(* IEC 61131-3 sources: SRCI_CLIENT_PLC/RobotLibrary/Library/Structures/AxesGroup/State/SyncState, 4 files *)

(* ---- AxesGroupStateSyncState.st ---- *)
{attribute 'pack_mode' := '1'}
// -------------------------------------------------------------------------
//  SRCI Robot Library
// -------------------------------------------------------------------------
//
//  Object:      AxesGroupStateSyncState
//  Author:      Thorsten Brach
//  Date:        2024-06-01
//
//  Description:
//
//
//  Copyright:
//    (C) 2024 Thorsten Brach. All rights reserved
//             Licensed under the MIT License.
//
//  Disclaimer:
//    This project is provided without any guarantee and can be used for
//    private and commercial purposes. Any use is at the user’s
//    own risk and responsibility.
//
// -------------------------------------------------------------------------
TYPE AxesGroupStateSyncState :
STRUCT
  /// Bit 00: Tool
  Tool             : BOOL;
  /// Bit 01: Frame
  Frame            : BOOL;
  /// Bit 02: Load
  Load             : BOOL;
  /// Bit 03: WorkArea
  WorkArea         : BOOL;
  /// Bit 04: SwLimits
  SwLimits         : BOOL;
  /// Bit 05: DefaultDynamics
  DefaultDynamics  : BOOL;
  /// Bit 06: ReferenceDynamics
  ReferenceDynamics: BOOL;
  /// Bit 07:
  Bit07            : BOOL;
  /// Bit 08:
  Bit08            : BOOL;
  /// Bit 09:
  Bit09            : BOOL;
  /// Bit 10:
  Bit10            : BOOL;
  /// Bit 11:
  Bit11            : BOOL;
  /// Bit 12:
  Bit12            : BOOL;
  /// Bit 13:
  Bit13            : BOOL;
  /// Bit 14:
  Bit14            : BOOL;
  /// Bit 15:
  Bit15            : BOOL;
END_STRUCT
END_TYPE

(* ---- AxesGroupStateSyncStateNo.st ---- *)
{attribute 'pack_mode' := '1'}
// -------------------------------------------------------------------------
//  SRCI Robot Library
// -------------------------------------------------------------------------
//
//  Object:      AxesGroupStateSyncStateNo
//  Author:      Thorsten Brach
//  Date:        2024-06-01
//
//  Description:
//
//
//  Copyright:
//    (C) 2024 Thorsten Brach. All rights reserved
//             Licensed under the MIT License.
//
//  Disclaimer:
//    This project is provided without any guarantee and can be used for
//    private and commercial purposes. Any use is at the user’s
//    own risk and responsibility.
//
// -------------------------------------------------------------------------
TYPE AxesGroupStateSyncStateNo :
STRUCT
  /// Ammount of unsynchronized tool data
  Tool     : USINT;
  /// Ammount of unsynchronized frame data
  Frame    : USINT;
  /// Ammount of unsynchronized load data
  Load     : USINT;
  /// Ammount of unsynchronized word areas
  WorkArea : USINT;
END_STRUCT
END_TYPE

(* ---- AxesGroupStateSyncStatePlc.st ---- *)
{attribute 'pack_mode' := '1'}
// -------------------------------------------------------------------------
//  SRCI Robot Library
// -------------------------------------------------------------------------
//
//  Object:      AxesGroupStateSyncStatePlc
//  Author:      Thorsten Brach
//  Date:        2024-06-01
//
//  Description:
//
//
//  Copyright:
//    (C) 2024 Thorsten Brach. All rights reserved
//             Licensed under the MIT License.
//
//  Disclaimer:
//    This project is provided without any guarantee and can be used for
//    private and commercial purposes. Any use is at the user’s
//    own risk and responsibility.
//
// -------------------------------------------------------------------------
TYPE AxesGroupStateSyncStatePlc :
STRUCT
  /// Synchronisation state of the datasets
  InSync   : AxesGroupStateSyncState;
  /// Number of the dataset which has been changed locally
  UnSyncNo : AxesGroupStateSyncStateNo;
END_STRUCT
END_TYPE

(* ---- AxesGroupStateSyncStateRob.st ---- *)
{attribute 'pack_mode' := '1'}
// -------------------------------------------------------------------------
//  SRCI Robot Library
// -------------------------------------------------------------------------
//
//  Object:      AxesGroupStateSyncStateRob
//  Author:      Thorsten Brach
//  Date:        2024-06-01
//
//  Description:
//
//
//  Copyright:
//    (C) 2024 Thorsten Brach. All rights reserved
//             Licensed under the MIT License.
//
//  Disclaimer:
//    This project is provided without any guarantee and can be used for
//    private and commercial purposes. Any use is at the user’s
//    own risk and responsibility.
//
// -------------------------------------------------------------------------
TYPE AxesGroupStateSyncStateRob :
STRUCT
  /// Synchronisation state of the datasets
  InSync   : AxesGroupStateSyncState;
  /// Number of the dataset which has been changed locally
  UnSyncNo : AxesGroupStateSyncStateNo;
END_STRUCT
END_TYPE
